// Mitsubishi GX Works2 project: Practica 2   PLC: FX3G

PROGRAM MAIN
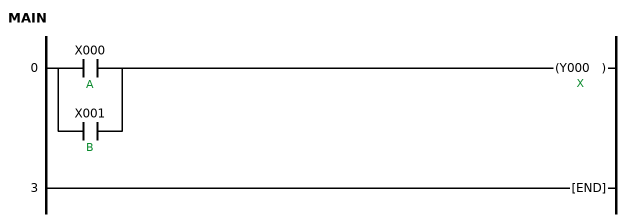
0     LD      X000  ; A
      OR      X001  ; B
      OUT     Y000  ; X
3     END
END_PROGRAM
